FUNCTION_BLOCK Atuador_Coester_HMI (* Service Interface Function Block Type *)
  (* Standard: 61499-2 *)
  (* Version 2.2, 04/11/2026, Hidryco, Hidryco, 2.2: STS_ALARME (IO List da Nereda). 2.1: restante das tags (posicao, torque, temperatura, tempo de percurso, status 2, alarmes), posicionar/parar so no posicionador, falha do atuador e faceplate de diagnostico. 2.0: refeito simples. *)
  PACKAGE Hidryco.HidrycoLib;
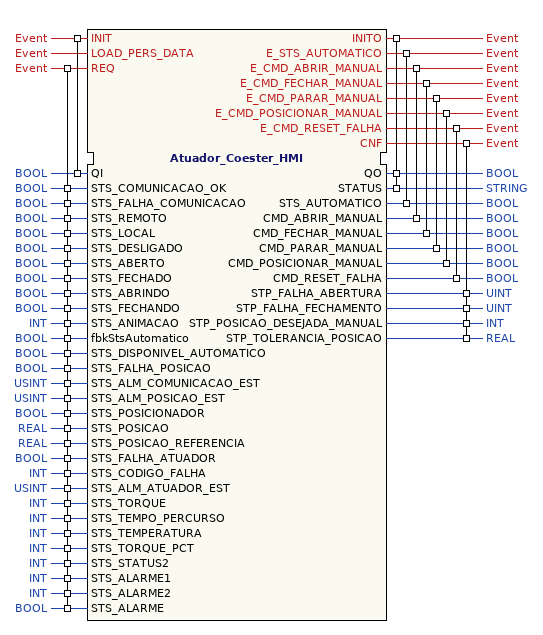
  EVENT_INPUT
    INIT WITH QI;
    LOAD_PERS_DATA; (* Reenvia os parametros persistentes *)
    REQ WITH STS_COMUNICACAO_OK, STS_FALHA_COMUNICACAO, STS_REMOTO, STS_LOCAL, STS_DESLIGADO, STS_ABERTO, STS_FECHADO, STS_ABRINDO, STS_FECHANDO, STS_ANIMACAO, fbkStsAutomatico, STS_DISPONIVEL_AUTOMATICO, STS_FALHA_POSICAO, STS_ALM_COMUNICACAO_EST, STS_ALM_POSICAO_EST, STS_POSICIONADOR, STS_POSICAO, STS_POSICAO_REFERENCIA, STS_FALHA_ATUADOR, STS_CODIGO_FALHA, STS_ALM_ATUADOR_EST, STS_TORQUE, STS_TEMPO_PERCURSO, STS_TEMPERATURA, STS_TORQUE_PCT, STS_STATUS2, STS_ALARME1, STS_ALARME2, STS_ALARME; (* Atualizacao de status *)
  END_EVENT
  EVENT_OUTPUT
    INITO WITH QO, STATUS;
    E_STS_AUTOMATICO WITH STS_AUTOMATICO;
    E_CMD_ABRIR_MANUAL WITH CMD_ABRIR_MANUAL;
    E_CMD_FECHAR_MANUAL WITH CMD_FECHAR_MANUAL;
    E_CMD_PARAR_MANUAL WITH CMD_PARAR_MANUAL;
    E_CMD_POSICIONAR_MANUAL WITH CMD_POSICIONAR_MANUAL;
    E_CMD_RESET_FALHA WITH CMD_RESET_FALHA;
    CNF WITH STP_FALHA_ABERTURA, STP_FALHA_FECHAMENTO, STP_POSICAO_DESEJADA_MANUAL, STP_TOLERANCIA_POSICAO;
  END_EVENT
  VAR_INPUT
    QI : BOOL;
    STS_COMUNICACAO_OK : BOOL; (* Comunicacao Modbus com o atuador OK *)
    STS_FALHA_COMUNICACAO : BOOL; (* Falha de comunicacao Modbus *)
    STS_REMOTO : BOOL; (* Seletor do atuador em Remoto *)
    STS_LOCAL : BOOL; (* Seletor do atuador em Local *)
    STS_DESLIGADO : BOOL; (* Seletor do atuador em Desligado *)
    STS_ABERTO : BOOL; (* Posicao aberta *)
    STS_FECHADO : BOOL; (* Posicao fechada *)
    STS_ABRINDO : BOOL; (* Em movimento de abertura *)
    STS_FECHANDO : BOOL; (* Em movimento de fechamento *)
    STS_ANIMACAO : INT; (* 0 fechada, 1 aberta, 2 falha, 3 intermediaria parada, 4 abrindo, 5 fechando *)
    fbkStsAutomatico : BOOL; (* Retorno do modo: TRUE = automatico *)
    STS_DISPONIVEL_AUTOMATICO : BOOL; (* Pode ser comandada pelo automatico agora *)
    STS_FALHA_POSICAO : BOOL; (* Nao abriu / nao fechou / nao posicionou no tempo (memorizada ate o reset) *)
    STS_ALM_COMUNICACAO_EST : USINT; (* Estado do ALARM_BIT comunicacao *)
    STS_ALM_POSICAO_EST : USINT; (* Estado do ALARM_BIT posicao *)
    STS_POSICIONADOR : BOOL; (* TRUE = instancia com posicionar e parar (cfgPosicionador) *)
    STS_POSICAO : REAL; (* Posicao real (%) - Word 5 *)
    STS_POSICAO_REFERENCIA : REAL; (* Ultima posicao enviada ao atuador (%) *)
    STS_FALHA_ATUADOR : BOOL; (* Falha do atuador (memorizada ate o reset) *)
    STS_CODIGO_FALHA : INT; (* Codigo da falha do atuador (texto na IHM) *)
    STS_ALM_ATUADOR_EST : USINT; (* Estado do ALARM_BIT falha do atuador *)
    STS_TORQUE : INT; (* Torque do ultimo comando (Nm) - Word 6 *)
    STS_TEMPO_PERCURSO : INT; (* Tempo do ultimo percurso (s) - Word 7 *)
    STS_TEMPERATURA : INT; (* Temperatura interna (graus C) - Word 8 - 19 *)
    STS_TORQUE_PCT : INT; (* Torque do ultimo comando (%) - Word 9 *)
    STS_STATUS2 : INT; (* Word 2 - status 2 *)
    STS_ALARME1 : INT; (* Word 3 - alarmes 1 *)
    STS_ALARME2 : INT; (* Word 4 - alarmes 2 *)
    STS_ALARME : BOOL; (* Alarme da valvula: falha de comunicacao OU falha do atuador OU nao abriu/fechou/posicionou *)
  END_VAR
  VAR_OUTPUT
    QO : BOOL; (* Event Output Qualifier *)
    STATUS : STRING; (* Service Status *)
    STS_AUTOMATICO : BOOL; (* Modo: TRUE = automatico (persistente; padrao automatico) *)
    CMD_ABRIR_MANUAL : BOOL; (* TRUE = abrir (manual) *)
    CMD_FECHAR_MANUAL : BOOL; (* TRUE = fechar (manual) *)
    CMD_PARAR_MANUAL : BOOL; (* TRUE = parar (manual, so posicionador) *)
    CMD_POSICIONAR_MANUAL : BOOL; (* TRUE = posicionar em STP_POSICAO_DESEJADA_MANUAL (so posicionador) *)
    CMD_RESET_FALHA : BOOL; (* Reset das falhas e reconhecimento dos alarmes *)
    STP_FALHA_ABERTURA : UINT; (* Tempo maximo para abrir/posicionar abrindo (s); 0 = sem supervisao *)
    STP_FALHA_FECHAMENTO : UINT; (* Tempo maximo para fechar/posicionar fechando (s); 0 = sem supervisao *)
    STP_POSICAO_DESEJADA_MANUAL : INT; (* Posicao desejada em manual (%) *)
    STP_TOLERANCIA_POSICAO : REAL; (* Tolerancia da posicao (%); 0 = 2 % *)
  END_VAR
  SERVICE /
    SEQUENCE 
    END_SEQUENCE
  END_SERVICE
END_FUNCTION_BLOCK
